Fanuc KAREL source: KC00063.KL

PROGRAM KC00063
%NOLOCKGROUP
%ENVIRONMENT CVIS
VAR
  I: INTEGER
  J: INTEGER
  K: INTEGER
  R: REAL
  B: BOOLEAN
  S: STRING[80]
  T: STRING[80]
  P: PATH
  Q: PATH
  AI: ARRAY[8] OF INTEGER
  AB: ARRAY[244] OF BYTE
BEGIN
  V_GET_QUEUE(I,J,K,I)
END KC00063
